KUKA KRL program: folge11.src, folge11.dat

--- folge11.src ---
&ACCESS RVP
&REL 1
&COMMENT bt2krl vw-ks24 production Folge 11 plan 16#F77E
DEF FOLGE11()
   ; Generated by bt2krl 0.1.0 from bt2plc plan bt_1790934549_welding_cell_2_small (cell welding_cell_2_small), PLAN_ID 16#F77E
   ; Robot robot1 (R1), controller 000001R01, model KR240R2900_ULTRA, joint mapping identity
   ; Profile vw-ks24 (VW KS24 / TPVW 8.1.8).
   ; Do not edit: regenerate with bt2krl (plain KRL, no inline forms).
   ; Production Folge: 8 ops; per op: op index BT_PKTNR, interlock request + MAKRO20 handshake, motion (exact stop at the end), hold, interlock release
   ; The VW tech package does the Folge handshake (cell.src, AUE_INIT/WAIT/END).
   ;FOLD AUE INIT
      VW(#VW_AUE_INIT,TRUE)
      PENTER:
      INTERRUPT DECL 10 WHEN $CYCFLAG[254]==FALSE DO VW(#FB_STOP,TRUE)
      INTERRUPT ON 10
      INT10=TRUE
   ;ENDFOLD
   ;FOLD VWP0 P0 10 PCT
      ; P0 = home: VW_INIT runs BAS(#INITMOV); AUE_WAIT later sets $H_POS here
      VW(#VW_INIT,TRUE)
      VW_USR_R (#USR_INIT)
      BAS(#VEL_PTP,10)
      $APO.CPTP=100
      PTP P0
      $OUT[15]=TRUE ; PF0 Grundstellung
      ; MAKRO0 RUECKSETZEN_EA: resets A33-A96 (also the tool releases)
      SEL_RES=SELECT(#MAKRO,0,TRUE,,,,,FALSE)
   ;ENDFOLD
   ;FOLD VWAUEWAIT
      VW(#VW_AUE_WAIT,TRUE )
      IF N_VW==TRUE THEN
         GOTO PEXIT
      ENDIF
   ;ENDFOLD
   ;FOLD VWSTART 16#00000003
      ; release every interlock this robot uses: IL01=V1 IL02=V11
      $OUT[15]=FALSE ; PF0 off
      ; MAKRO50 Ini Merker: the cyclic flags of the driving conditions
      SEL_RES=SELECT(#MAKRO,50,TRUE,,,,,FALSE)
      $OUT[41]=TRUE ; release V1
      $OUT[51]=TRUE ; release V11
   ;ENDFOLD
   ;FOLD PLAN ID 16#F77E
      IF BT_PLANID<>PLAN_ID THEN
         $LOOP_MSG[]="BT2KRL PLAN_ID mismatch - regenerate KRL and PLC"
         HALT
      ENDIF
   ;ENDFOLD
   ;FOLD VWFB 16#00000000
      VALCYCFL30=$CYCFLAG[254]
      $CYCFLAG[254]=($CYCFLAG[30]) AND $CYCFLAG[255] OR ($TIMER[61]<0)
      VW(#FB_CHECK,TRUE)
   ;ENDFOLD
   ;FOLD OP 1 W01 MASK 16#00000001
      ; zones IL01
      BT_PKTNR=1
      ;FOLD VWLOCK 16#00000001
         ; enter IL01=V1
         $OUT[81]=TRUE ; request V1
         ; MAKRO20 semantics, inline for these interlocks only
         $OUT[41]=$OUT[41] OR $OUT[81]
         ; PLC grant of the request
         $LOOP_MSG[]="E81"
         $LOOP_CONT=TRUE
         WAIT FOR ($IN[81]) OR (NOT $LOOP_CONT AND ($MODE_OP<>#EX))
         $LOOP_MSG[]="                                                                                                                                "
         ; partner release
         $LOOP_MSG[]="E41"
         $LOOP_CONT=TRUE
         WAIT FOR ($IN[41]) OR (NOT $LOOP_CONT AND ($MODE_OP<>#EX))
         $LOOP_MSG[]="                                                                                                                                "
         $OUT[41]=FALSE ; occupied
         $OUT[81]=FALSE
      ;ENDFOLD
      ;FOLD VWFB 16#00000001
         VALCYCFL30=$CYCFLAG[254]
         $CYCFLAG[254]=($CYCFLAG[30] AND $IN[41]) AND $CYCFLAG[255] OR ($TIMER[61]<0)
         VW(#FB_CHECK,TRUE)
      ;ENDFOLD
      BAS(#VEL_PTP,3)
      PTP P1 C_PTP
      BAS(#VEL_PTP,6)
      PTP P2 C_PTP
      BAS(#VEL_PTP,10)
      PTP P3 C_PTP
      BAS(#VEL_PTP,12)
      PTP P4 C_PTP
      BAS(#VEL_PTP,15)
      PTP P5 C_PTP
      BAS(#VEL_PTP,17)
      PTP P6 C_PTP
      BAS(#VEL_PTP,19)
      PTP P7 C_PTP
      BAS(#VEL_PTP,17)
      PTP P8 C_PTP
      BAS(#VEL_PTP,13)
      PTP P9 C_PTP
      BAS(#VEL_PTP,10)
      PTP P10 C_PTP
      BAS(#VEL_PTP,6)
      PTP P11 C_PTP
      BAS(#VEL_PTP,3)
      PTP P12 C_PTP
      BAS(#VEL_PTP,5)
      PTP P13 C_PTP
      BAS(#VEL_PTP,4)
      PTP P14
      WAIT SEC 0.5 ; hold
      ;FOLD VWUNLOCK 16#00000001
         ; leave IL01=V1
         $OUT[41]=TRUE ; release V1
      ;ENDFOLD
      ;FOLD VWFB 16#00000000
         VALCYCFL30=$CYCFLAG[254]
         $CYCFLAG[254]=($CYCFLAG[30]) AND $CYCFLAG[255] OR ($TIMER[61]<0)
         VW(#FB_CHECK,TRUE)
      ;ENDFOLD
      WAIT SEC 0.1 ; step dwell
   ;ENDFOLD
   ;FOLD OP 2 W02 MASK 16#00000002
      ; zones IL02
      BT_PKTNR=2
      ;FOLD VWLOCK 16#00000002
         ; enter IL02=V11
         $OUT[91]=TRUE ; request V11
         ; MAKRO20 semantics, inline for these interlocks only
         $OUT[51]=$OUT[51] OR $OUT[91]
         ; PLC grant of the request
         $LOOP_MSG[]="E91"
         $LOOP_CONT=TRUE
         WAIT FOR ($IN[91]) OR (NOT $LOOP_CONT AND ($MODE_OP<>#EX))
         $LOOP_MSG[]="                                                                                                                                "
         ; partner release
         $LOOP_MSG[]="E51"
         $LOOP_CONT=TRUE
         WAIT FOR ($IN[51]) OR (NOT $LOOP_CONT AND ($MODE_OP<>#EX))
         $LOOP_MSG[]="                                                                                                                                "
         $OUT[51]=FALSE ; occupied
         $OUT[91]=FALSE
      ;ENDFOLD
      ;FOLD VWFB 16#00000002
         VALCYCFL30=$CYCFLAG[254]
         $CYCFLAG[254]=($CYCFLAG[30] AND $IN[51]) AND $CYCFLAG[255] OR ($TIMER[61]<0)
         VW(#FB_CHECK,TRUE)
      ;ENDFOLD
      BAS(#VEL_PTP,3)
      PTP P15 C_PTP
      BAS(#VEL_PTP,7)
      PTP P16 C_PTP
      BAS(#VEL_PTP,10)
      PTP P17 C_PTP
      BAS(#VEL_PTP,13)
      PTP P18 C_PTP
      BAS(#VEL_PTP,10)
      PTP P19 C_PTP
      BAS(#VEL_PTP,7)
      PTP P20 C_PTP
      BAS(#VEL_PTP,3)
      PTP P21 C_PTP
      BAS(#VEL_PTP,5)
      PTP P22 C_PTP
      BAS(#VEL_PTP,4)
      PTP P23
      WAIT SEC 0.5 ; hold
      ;FOLD VWUNLOCK 16#00000002
         ; leave IL02=V11
         $OUT[51]=TRUE ; release V11
      ;ENDFOLD
      ;FOLD VWFB 16#00000000
         VALCYCFL30=$CYCFLAG[254]
         $CYCFLAG[254]=($CYCFLAG[30]) AND $CYCFLAG[255] OR ($TIMER[61]<0)
         VW(#FB_CHECK,TRUE)
      ;ENDFOLD
      WAIT SEC 0.1 ; step dwell
   ;ENDFOLD
   ;FOLD OP 3 W03 MASK 16#00000001
      ; zones IL01
      BT_PKTNR=3
      ;FOLD VWLOCK 16#00000001
         ; enter IL01=V1
         $OUT[81]=TRUE ; request V1
         ; MAKRO20 semantics, inline for these interlocks only
         $OUT[41]=$OUT[41] OR $OUT[81]
         ; PLC grant of the request
         $LOOP_MSG[]="E81"
         $LOOP_CONT=TRUE
         WAIT FOR ($IN[81]) OR (NOT $LOOP_CONT AND ($MODE_OP<>#EX))
         $LOOP_MSG[]="                                                                                                                                "
         ; partner release
         $LOOP_MSG[]="E41"
         $LOOP_CONT=TRUE
         WAIT FOR ($IN[41]) OR (NOT $LOOP_CONT AND ($MODE_OP<>#EX))
         $LOOP_MSG[]="                                                                                                                                "
         $OUT[41]=FALSE ; occupied
         $OUT[81]=FALSE
      ;ENDFOLD
      ;FOLD VWFB 16#00000001
         VALCYCFL30=$CYCFLAG[254]
         $CYCFLAG[254]=($CYCFLAG[30] AND $IN[41]) AND $CYCFLAG[255] OR ($TIMER[61]<0)
         VW(#FB_CHECK,TRUE)
      ;ENDFOLD
      BAS(#VEL_PTP,2)
      PTP P24 C_PTP
      BAS(#VEL_PTP,6)
      PTP P25 C_PTP
      BAS(#VEL_PTP,9)
      PTP P26 C_PTP
      BAS(#VEL_PTP,13)
      PTP P27 C_PTP
      BAS(#VEL_PTP,15)
      PTP P28 C_PTP
      BAS(#VEL_PTP,12)
      PTP P29 C_PTP
      BAS(#VEL_PTP,8)
      PTP P30 C_PTP
      BAS(#VEL_PTP,6)
      PTP P31 C_PTP
      BAS(#VEL_PTP,2)
      PTP P32 C_PTP
      BAS(#VEL_PTP,6)
      PTP P33 C_PTP
      BAS(#VEL_PTP,8)
      PTP P34 C_PTP
      BAS(#VEL_PTP,4)
      PTP P35
      WAIT SEC 0.5 ; hold
      ;FOLD VWUNLOCK 16#00000001
         ; leave IL01=V1
         $OUT[41]=TRUE ; release V1
      ;ENDFOLD
      ;FOLD VWFB 16#00000000
         VALCYCFL30=$CYCFLAG[254]
         $CYCFLAG[254]=($CYCFLAG[30]) AND $CYCFLAG[255] OR ($TIMER[61]<0)
         VW(#FB_CHECK,TRUE)
      ;ENDFOLD
      WAIT SEC 0.1 ; step dwell
   ;ENDFOLD
   ;FOLD OP 4 W06 MASK 16#00000002
      ; zones IL02
      BT_PKTNR=4
      ;FOLD VWLOCK 16#00000002
         ; enter IL02=V11
         $OUT[91]=TRUE ; request V11
         ; MAKRO20 semantics, inline for these interlocks only
         $OUT[51]=$OUT[51] OR $OUT[91]
         ; PLC grant of the request
         $LOOP_MSG[]="E91"
         $LOOP_CONT=TRUE
         WAIT FOR ($IN[91]) OR (NOT $LOOP_CONT AND ($MODE_OP<>#EX))
         $LOOP_MSG[]="                                                                                                                                "
         ; partner release
         $LOOP_MSG[]="E51"
         $LOOP_CONT=TRUE
         WAIT FOR ($IN[51]) OR (NOT $LOOP_CONT AND ($MODE_OP<>#EX))
         $LOOP_MSG[]="                                                                                                                                "
         $OUT[51]=FALSE ; occupied
         $OUT[91]=FALSE
      ;ENDFOLD
      ;FOLD VWFB 16#00000002
         VALCYCFL30=$CYCFLAG[254]
         $CYCFLAG[254]=($CYCFLAG[30] AND $IN[51]) AND $CYCFLAG[255] OR ($TIMER[61]<0)
         VW(#FB_CHECK,TRUE)
      ;ENDFOLD
      BAS(#VEL_PTP,8)
      PTP P36 C_PTP
      BAS(#VEL_PTP,16)
      PTP P37 C_PTP
      BAS(#VEL_PTP,8)
      PTP P38 C_PTP
      BAS(#VEL_PTP,4)
      PTP P39 C_PTP
      BAS(#VEL_PTP,3)
      PTP P40
      WAIT SEC 0.5 ; hold
      ;FOLD VWUNLOCK 16#00000002
         ; leave IL02=V11
         $OUT[51]=TRUE ; release V11
      ;ENDFOLD
      ;FOLD VWFB 16#00000000
         VALCYCFL30=$CYCFLAG[254]
         $CYCFLAG[254]=($CYCFLAG[30]) AND $CYCFLAG[255] OR ($TIMER[61]<0)
         VW(#FB_CHECK,TRUE)
      ;ENDFOLD
      WAIT SEC 0.1 ; step dwell
   ;ENDFOLD
   ;FOLD OP 5 W05 MASK 16#00000001
      ; zones IL01
      BT_PKTNR=5
      ;FOLD VWLOCK 16#00000001
         ; enter IL01=V1
         $OUT[81]=TRUE ; request V1
         ; MAKRO20 semantics, inline for these interlocks only
         $OUT[41]=$OUT[41] OR $OUT[81]
         ; PLC grant of the request
         $LOOP_MSG[]="E81"
         $LOOP_CONT=TRUE
         WAIT FOR ($IN[81]) OR (NOT $LOOP_CONT AND ($MODE_OP<>#EX))
         $LOOP_MSG[]="                                                                                                                                "
         ; partner release
         $LOOP_MSG[]="E41"
         $LOOP_CONT=TRUE
         WAIT FOR ($IN[41]) OR (NOT $LOOP_CONT AND ($MODE_OP<>#EX))
         $LOOP_MSG[]="                                                                                                                                "
         $OUT[41]=FALSE ; occupied
         $OUT[81]=FALSE
      ;ENDFOLD
      ;FOLD VWFB 16#00000001
         VALCYCFL30=$CYCFLAG[254]
         $CYCFLAG[254]=($CYCFLAG[30] AND $IN[41]) AND $CYCFLAG[255] OR ($TIMER[61]<0)
         VW(#FB_CHECK,TRUE)
      ;ENDFOLD
      BAS(#VEL_PTP,2)
      PTP P41 C_PTP
      BAS(#VEL_PTP,6)
      PTP P42 C_PTP
      BAS(#VEL_PTP,10)
      PTP P43 C_PTP
      BAS(#VEL_PTP,13)
      PTP P44 C_PTP
      BAS(#VEL_PTP,15)
      PTP P45 C_PTP
      BAS(#VEL_PTP,12)
      PTP P46 C_PTP
      BAS(#VEL_PTP,8)
      PTP P47 C_PTP
      BAS(#VEL_PTP,6)
      PTP P48 C_PTP
      BAS(#VEL_PTP,2)
      PTP P49 C_PTP
      BAS(#VEL_PTP,4)
      PTP P50 C_PTP
      PTP P51
      WAIT SEC 0.5 ; hold
      ;FOLD VWUNLOCK 16#00000001
         ; leave IL01=V1
         $OUT[41]=TRUE ; release V1
      ;ENDFOLD
      ;FOLD VWFB 16#00000000
         VALCYCFL30=$CYCFLAG[254]
         $CYCFLAG[254]=($CYCFLAG[30]) AND $CYCFLAG[255] OR ($TIMER[61]<0)
         VW(#FB_CHECK,TRUE)
      ;ENDFOLD
      WAIT SEC 0.1 ; step dwell
   ;ENDFOLD
   ;FOLD OP 6 W04 MASK 16#00000002
      ; zones IL02
      BT_PKTNR=6
      ;FOLD VWLOCK 16#00000002
         ; enter IL02=V11
         $OUT[91]=TRUE ; request V11
         ; MAKRO20 semantics, inline for these interlocks only
         $OUT[51]=$OUT[51] OR $OUT[91]
         ; PLC grant of the request
         $LOOP_MSG[]="E91"
         $LOOP_CONT=TRUE
         WAIT FOR ($IN[91]) OR (NOT $LOOP_CONT AND ($MODE_OP<>#EX))
         $LOOP_MSG[]="                                                                                                                                "
         ; partner release
         $LOOP_MSG[]="E51"
         $LOOP_CONT=TRUE
         WAIT FOR ($IN[51]) OR (NOT $LOOP_CONT AND ($MODE_OP<>#EX))
         $LOOP_MSG[]="                                                                                                                                "
         $OUT[51]=FALSE ; occupied
         $OUT[91]=FALSE
      ;ENDFOLD
      ;FOLD VWFB 16#00000002
         VALCYCFL30=$CYCFLAG[254]
         $CYCFLAG[254]=($CYCFLAG[30] AND $IN[51]) AND $CYCFLAG[255] OR ($TIMER[61]<0)
         VW(#FB_CHECK,TRUE)
      ;ENDFOLD
      BAS(#VEL_PTP,3)
      PTP P52 C_PTP
      BAS(#VEL_PTP,7)
      PTP P53 C_PTP
      BAS(#VEL_PTP,10)
      PTP P54 C_PTP
      BAS(#VEL_PTP,13)
      PTP P55 C_PTP
      BAS(#VEL_PTP,11)
      PTP P56 C_PTP
      BAS(#VEL_PTP,7)
      PTP P57 C_PTP
      BAS(#VEL_PTP,3)
      PTP P58 C_PTP
      BAS(#VEL_PTP,4)
      PTP P59 C_PTP
      BAS(#VEL_PTP,3)
      PTP P60
      WAIT SEC 0.5 ; hold
      ;FOLD VWUNLOCK 16#00000002
         ; leave IL02=V11
         $OUT[51]=TRUE ; release V11
      ;ENDFOLD
      ;FOLD VWFB 16#00000000
         VALCYCFL30=$CYCFLAG[254]
         $CYCFLAG[254]=($CYCFLAG[30]) AND $CYCFLAG[255] OR ($TIMER[61]<0)
         VW(#FB_CHECK,TRUE)
      ;ENDFOLD
      WAIT SEC 0.1 ; step dwell
   ;ENDFOLD
   ;FOLD OP 7 R1_PARK MASK 16#00000001
      ; zones IL01
      BT_PKTNR=7
      ;FOLD VWLOCK 16#00000001
         ; enter IL01=V1
         $OUT[81]=TRUE ; request V1
         ; MAKRO20 semantics, inline for these interlocks only
         $OUT[41]=$OUT[41] OR $OUT[81]
         ; PLC grant of the request
         $LOOP_MSG[]="E81"
         $LOOP_CONT=TRUE
         WAIT FOR ($IN[81]) OR (NOT $LOOP_CONT AND ($MODE_OP<>#EX))
         $LOOP_MSG[]="                                                                                                                                "
         ; partner release
         $LOOP_MSG[]="E41"
         $LOOP_CONT=TRUE
         WAIT FOR ($IN[41]) OR (NOT $LOOP_CONT AND ($MODE_OP<>#EX))
         $LOOP_MSG[]="                                                                                                                                "
         $OUT[41]=FALSE ; occupied
         $OUT[81]=FALSE
      ;ENDFOLD
      ;FOLD VWFB 16#00000001
         VALCYCFL30=$CYCFLAG[254]
         $CYCFLAG[254]=($CYCFLAG[30] AND $IN[41]) AND $CYCFLAG[255] OR ($TIMER[61]<0)
         VW(#FB_CHECK,TRUE)
      ;ENDFOLD
      BAS(#VEL_PTP,6)
      PTP P61 C_PTP
      BAS(#VEL_PTP,14)
      PTP P62 C_PTP
      BAS(#VEL_PTP,22)
      PTP P63 C_PTP
      BAS(#VEL_PTP,19)
      PTP P64 C_PTP
      BAS(#VEL_PTP,13)
      PTP P65 C_PTP
      BAS(#VEL_PTP,25)
      PTP P66 C_PTP
      PTP P67
      WAIT SEC 0.5 ; hold
      ;FOLD VWUNLOCK 16#00000001
         ; leave IL01=V1
         $OUT[41]=TRUE ; release V1
      ;ENDFOLD
      ;FOLD VWFB 16#00000000
         VALCYCFL30=$CYCFLAG[254]
         $CYCFLAG[254]=($CYCFLAG[30]) AND $CYCFLAG[255] OR ($TIMER[61]<0)
         VW(#FB_CHECK,TRUE)
      ;ENDFOLD
      WAIT SEC 0.1 ; step dwell
   ;ENDFOLD
   ;FOLD OP 8 HOME MASK 16#00000002
      ; zones IL02
      BT_PKTNR=8
      ;FOLD VWLOCK 16#00000002
         ; enter IL02=V11
         $OUT[91]=TRUE ; request V11
         ; MAKRO20 semantics, inline for these interlocks only
         $OUT[51]=$OUT[51] OR $OUT[91]
         ; PLC grant of the request
         $LOOP_MSG[]="E91"
         $LOOP_CONT=TRUE
         WAIT FOR ($IN[91]) OR (NOT $LOOP_CONT AND ($MODE_OP<>#EX))
         $LOOP_MSG[]="                                                                                                                                "
         ; partner release
         $LOOP_MSG[]="E51"
         $LOOP_CONT=TRUE
         WAIT FOR ($IN[51]) OR (NOT $LOOP_CONT AND ($MODE_OP<>#EX))
         $LOOP_MSG[]="                                                                                                                                "
         $OUT[51]=FALSE ; occupied
         $OUT[91]=FALSE
      ;ENDFOLD
      ;FOLD VWFB 16#00000002
         VALCYCFL30=$CYCFLAG[254]
         $CYCFLAG[254]=($CYCFLAG[30] AND $IN[51]) AND $CYCFLAG[255] OR ($TIMER[61]<0)
         VW(#FB_CHECK,TRUE)
      ;ENDFOLD
      BAS(#VEL_PTP,3)
      PTP P68 C_PTP
      BAS(#VEL_PTP,8)
      PTP P69 C_PTP
      BAS(#VEL_PTP,12)
      PTP P70 C_PTP
      BAS(#VEL_PTP,17)
      PTP P71 C_PTP
      BAS(#VEL_PTP,20)
      PTP P72 C_PTP
      BAS(#VEL_PTP,23)
      PTP P73 C_PTP
      BAS(#VEL_PTP,26)
      PTP P74 C_PTP
      BAS(#VEL_PTP,27)
      PTP P75 C_PTP
      BAS(#VEL_PTP,24)
      PTP P76 C_PTP
      BAS(#VEL_PTP,22)
      PTP P77 C_PTP
      BAS(#VEL_PTP,18)
      PTP P78 C_PTP
      BAS(#VEL_PTP,14)
      PTP P79 C_PTP
      BAS(#VEL_PTP,9)
      PTP P80 C_PTP
      BAS(#VEL_PTP,3)
      PTP P81
      ;FOLD VWMAKRO 15
         ; Gesamtfertigmeldung
         SEL_RES=SELECT(#MAKRO,15,TRUE,,,,,FALSE)
      ;ENDFOLD
      ;FOLD VWUNLOCK 16#00000002
         ; leave IL02=V11
         $OUT[51]=TRUE ; release V11
      ;ENDFOLD
      ;FOLD VWFB 16#00000000
         VALCYCFL30=$CYCFLAG[254]
         $CYCFLAG[254]=($CYCFLAG[30]) AND $CYCFLAG[255] OR ($TIMER[61]<0)
         VW(#FB_CHECK,TRUE)
      ;ENDFOLD
      WAIT SEC 0.1 ; step dwell
   ;ENDFOLD
   BT_PKTNR=0
   ;FOLD AUE END
      VW(#VW_AUE_END,TRUE)
      GOTO PENTER
      PEXIT:
   ;ENDFOLD
END

--- folge11.dat ---
&ACCESS RVP
&REL 1
&COMMENT bt2krl vw-ks24 data Folge 11 plan 16#F77E
DEFDAT FOLGE11
   ; Generated by bt2krl 0.1.0 from bt2plc plan bt_1790934549_welding_cell_2_small (cell welding_cell_2_small), PLAN_ID 16#F77E
   ; Robot robot1 (R1), controller 000001R01, model KR240R2900_ULTRA, joint mapping identity
   ; Profile vw-ks24 (VW KS24 / TPVW 8.1.8).
   ; Do not edit: regenerate with bt2krl (plain KRL, no inline forms).
   EXT BAS (BAS_COMMAND :IN,REAL :IN )
   ; interface to the VW standard routines (as every VW Folge .dat declares them)
   EXT VW (VW_COMMAND :IN,BOOL :IN,REAL :IN,REAL :IN,REAL :IN,REAL :IN,BOOL :IN,E6POS :IN )
   EXT VW_USR_R (VW_USER_CMD :IN,INT :IN,REAL :IN,REAL :IN,REAL :IN,REAL :IN,REAL :IN,REAL :IN,BOOL :IN )
   EXTFCT INT SELECT (SUBTYPE :IN,INT :IN,BOOL :IN,ARI_TYP :IN,INT :IN,BOOL_TYP :IN,INT :IN,BOOL :IN)
   DECL AXIS P0={A1 0.0,A2 -90.0,A3 90.0,A4 0.0,A5 0.0,A6 0.0}
   DECL AXIS P1={A1 -1.1481,A2 -89.8273,A3 90.1392,A4 0.2955,A5 0.7752,A6 0.3515}
   DECL AXIS P2={A1 -4.4157,A2 -89.3356,A3 90.5354,A4 1.1366,A5 2.9817,A6 1.3518}
   DECL AXIS P3={A1 -9.5379,A2 -88.565,A3 91.1564,A4 2.455,A5 6.4405,A6 2.9199}
   DECL AXIS P4={A1 -16.2497,A2 -87.5551,A3 91.9702,A4 4.1827,A5 10.9727,A6 4.9746}
   DECL AXIS P5={A1 -24.2863,A2 -86.346,A3 92.9446,A4 6.2512,A5 16.3994,A6 7.4349}
   DECL AXIS P6={A1 -38.2454,A2 -84.2458,A3 94.6371,A4 9.8443,A5 25.8253,A6 11.7083}
   DECL AXIS P7={A1 -90.5161,A2 -76.3814,A3 100.9747,A4 23.2987,A5 61.1212,A6 27.7103}
   DECL AXIS P8={A1 -108.6425,A2 -73.6542,A3 103.1724,A4 27.9644,A5 73.3611,A6 33.2594}
   DECL AXIS P9={A1 -119.2236,A2 -72.0622,A3 104.4553,A4 30.6879,A5 80.506,A6 36.4987}
   DECL AXIS P10={A1 -124.3458,A2 -71.2916,A3 105.0764,A4 32.0064,A5 83.9648,A6 38.0668}
   DECL AXIS P11={A1 -127.6134,A2 -70.7999,A3 105.4725,A4 32.8474,A5 86.1712,A6 39.0671}
   DECL AXIS P12={A1 -128.7615,A2 -70.6272,A3 105.6117,A4 33.143,A5 86.9465,A6 39.4186}
   DECL AXIS P13={A1 -128.7615,A2 -70.2228,A3 105.9156,A4 33.18,A5 86.8872,A6 39.3731}
   DECL AXIS P14={A1 -128.7615,A2 -67.4517,A3 107.7396,A4 33.6697,A5 83.7898,A6 37.2493}
   DECL AXIS P15={A1 -128.6426,A2 -67.6366,A3 107.8186,A4 32.7502,A5 82.9536,A6 37.7433}
   DECL AXIS P16={A1 -128.3199,A2 -68.1386,A3 108.0329,A4 30.2544,A5 80.6837,A6 39.084}
   DECL AXIS P17={A1 -127.8443,A2 -68.8784,A3 108.3488,A4 26.5764,A5 77.3387,A6 41.0597}
   DECL AXIS P18={A1 -125.4325,A2 -72.6301,A3 109.9508,A4 7.9238,A5 60.3747,A6 51.0796}
   DECL AXIS P19={A1 -124.957,A2 -73.3699,A3 110.2667,A4 4.2458,A5 57.0297,A6 53.0553}
   DECL AXIS P20={A1 -124.6342,A2 -73.8718,A3 110.481,A4 1.75,A5 54.7598,A6 54.396}
   DECL AXIS P21={A1 -124.5154,A2 -74.0568,A3 110.56,A4 0.8305,A5 53.9236,A6 54.8899}
   DECL AXIS P22={A1 -124.5151,A2 -73.6213,A3 110.8768,A4 0.5687,A5 53.3206,A6 55.0767}
   DECL AXIS P23={A1 -124.5148,A2 -70.6583,A3 112.7632,A4 0.0121,A5 48.729,A6 55.4761}
   DECL AXIS P24={A1 -124.4617,A2 -70.7313,A3 112.7862,A4 -0.6572,A5 48.6812,A6 55.9965}
   DECL AXIS P25={A1 -124.3117,A2 -70.9378,A3 112.8512,A4 -2.5487,A5 48.5461,A6 57.4671}
   DECL AXIS P26={A1 -123.7762,A2 -71.6746,A3 113.0835,A4 -9.2998,A5 48.0639,A6 62.7161}
   DECL AXIS P27={A1 -123.0192,A2 -72.7163,A3 113.4118,A4 -18.8444,A5 47.3821,A6 70.1371}
   DECL AXIS P28={A1 -120.8842,A2 -75.654,A3 114.3378,A4 -45.7616,A5 45.4595,A6 91.0652}
   DECL AXIS P29={A1 -120.2241,A2 -76.5623,A3 114.6241,A4 -54.084,A5 44.865,A6 97.536}
   DECL AXIS P30={A1 -119.991,A2 -76.883,A3 114.7252,A4 -57.0231,A5 44.6551,A6 99.8211}
   DECL AXIS P31={A1 -119.8409,A2 -77.0895,A3 114.7902,A4 -58.9146,A5 44.52,A6 101.2917}
   DECL AXIS P32={A1 -119.7879,A2 -77.1625,A3 114.8133,A4 -59.5839,A5 44.4722,A6 101.8121}
   DECL AXIS P33={A1 -119.7876,A2 -76.7001,A3 115.1416,A4 -60.3559,A5 44.324,A6 102.6809}
   DECL AXIS P34={A1 -119.7872,A2 -76.0201,A3 115.6192,A4 -61.4852,A5 44.0795,A6 103.9753}
   DECL AXIS P35={A1 -119.7872,A2 -73.5459,A3 117.1,A4 -65.4365,A5 42.4249,A6 109.2463}
   DECL AXIS P36={A1 -119.1489,A2 -72.8001,A3 114.8711,A4 -64.2164,A5 43.4199,A6 108.0229}
   DECL AXIS P37={A1 -116.34,A2 -69.5185,A3 105.0638,A4 -58.8479,A5 47.7981,A6 102.6395}
   DECL AXIS P38={A1 -115.7016,A2 -68.7727,A3 102.8349,A4 -57.6278,A5 48.7931,A6 101.416}
   DECL AXIS P39={A1 -115.7012,A2 -68.3831,A3 103.1319,A4 -57.6419,A5 48.7925,A6 101.457}
   DECL AXIS P40={A1 -115.7007,A2 -65.7101,A3 104.9261,A4 -60.3105,A5 47.1665,A6 105.7542}
   DECL AXIS P41={A1 -115.7494,A2 -65.7146,A3 104.8564,A4 -59.6416,A5 47.2762,A6 105.2455}
   DECL AXIS P42={A1 -115.887,A2 -65.727,A3 104.6592,A4 -57.7513,A5 47.5859,A6 103.8079}
   DECL AXIS P43={A1 -116.378,A2 -65.7715,A3 103.9556,A4 -51.0043,A5 48.6915,A6 98.6766}
   DECL AXIS P44={A1 -117.0722,A2 -65.8345,A3 102.9609,A4 -41.4655,A5 50.2545,A6 91.4221}
   DECL AXIS P45={A1 -119.0301,A2 -66.012,A3 100.1555,A4 -14.5649,A5 54.6625,A6 70.9633}
   DECL AXIS P46={A1 -119.6354,A2 -66.0668,A3 99.2881,A4 -6.2475,A5 56.0254,A6 64.6377}
   DECL AXIS P47={A1 -119.8492,A2 -66.0862,A3 98.9818,A4 -3.3103,A5 56.5068,A6 62.4038}
   DECL AXIS P48={A1 -119.9868,A2 -66.0987,A3 98.7847,A4 -1.42,A5 56.8165,A6 60.9662}
   DECL AXIS P49={A1 -120.0355,A2 -66.1031,A3 98.7149,A4 -0.7511,A5 56.9261,A6 60.4575}
   DECL AXIS P50={A1 -120.0357,A2 -65.7312,A3 99.0104,A4 -0.6308,A5 56.7548,A6 60.3791}
   DECL AXIS P51={A1 -120.0359,A2 -63.1985,A3 100.772,A4 -0.0303,A5 53.2125,A6 59.9847}
   DECL AXIS P52={A1 -120.1288,A2 -63.1954,A3 100.6111,A4 0.7952,A5 54.0248,A6 59.6456}
   DECL AXIS P53={A1 -120.3834,A2 -63.1866,A3 100.1699,A4 3.0584,A5 56.2523,A6 58.7158}
   DECL AXIS P54={A1 -120.7638,A2 -63.1736,A3 99.5107,A4 6.44,A5 59.5803,A6 57.3266}
   DECL AXIS P55={A1 -122.8245,A2 -63.1028,A3 95.9394,A4 24.7593,A5 77.6095,A6 49.8008}
   DECL AXIS P56={A1 -123.6751,A2 -63.0736,A3 94.4653,A4 32.3213,A5 85.0518,A6 46.6942}
   DECL AXIS P57={A1 -123.9297,A2 -63.0649,A3 94.024,A4 34.5845,A5 87.2792,A6 45.7644}
   DECL AXIS P58={A1 -124.0225,A2 -63.0617,A3 93.8631,A4 35.41,A5 88.0916,A6 45.4253}
   DECL AXIS P59={A1 -124.0227,A2 -62.712,A3 94.1541,A4 35.4756,A5 88.0225,A6 45.3131}
   DECL AXIS P60={A1 -124.0229,A2 -60.325,A3 95.8907,A4 35.9822,A5 85.4859,A6 43.0775}
   DECL AXIS P61={A1 -125.6247,A2 -60.4541,A3 95.8014,A4 35.9822,A5 85.4859,A6 43.0775}
   DECL AXIS P62={A1 -129.8294,A2 -60.7871,A3 95.5713,A4 35.9822,A5 85.4859,A6 43.0775}
   DECL AXIS P63={A1 -149.0509,A2 -62.195,A3 94.602,A4 35.9822,A5 85.4859,A6 43.0775}
   DECL AXIS P64={A1 -154.6572,A2 -62.529,A3 94.3745,A4 35.9822,A5 85.4859,A6 43.0775}
   DECL AXIS P65={A1 -158.3613,A2 -62.6594,A3 94.2891,A4 35.9822,A5 85.4859,A6 43.0775}
   DECL AXIS P66={A1 -160.5075,A2 -61.5043,A3 95.1253,A4 35.9822,A5 85.4859,A6 43.0775}
   DECL AXIS P67={A1 -158.3613,A2 -60.3464,A3 95.9536,A4 35.9822,A5 85.4859,A6 43.0775}
   DECL AXIS P68={A1 -157.2676,A2 -60.5512,A3 95.9125,A4 35.7336,A5 84.8955,A6 42.78}
   DECL AXIS P69={A1 -154.1335,A2 -61.1381,A3 95.7947,A4 35.0215,A5 83.2037,A6 41.9274}
   DECL AXIS P70={A1 -149.1796,A2 -62.0657,A3 95.6084,A4 33.8959,A5 80.5295,A6 40.5799}
   DECL AXIS P71={A1 -138.8192,A2 -64.0057,A3 95.2189,A4 31.5419,A5 74.9368,A6 37.7616}
   DECL AXIS P72={A1 -130.2809,A2 -65.6046,A3 94.8979,A4 29.6018,A5 70.3276,A6 35.439}
   DECL AXIS P73={A1 -115.5777,A2 -68.3578,A3 94.3452,A4 26.2611,A5 62.3907,A6 31.4395}
   DECL AXIS P74={A1 -99.2616,A2 -71.413,A3 93.7317,A4 22.5538,A5 53.583,A6 27.0012}
   DECL AXIS P75={A1 -48.0798,A2 -80.9969,A3 91.8076,A4 10.9245,A5 25.9542,A6 13.0787}
   DECL AXIS P76={A1 -32.7563,A2 -83.8663,A3 91.2315,A4 7.4427,A5 17.6824,A6 8.9104}
   DECL AXIS P77={A1 -23.6665,A2 -85.5684,A3 90.8897,A4 5.3774,A5 12.7756,A6 6.4378}
   DECL AXIS P78={A1 -12.2721,A2 -87.702,A3 90.4614,A4 2.7884,A5 6.6247,A6 3.3383}
   DECL AXIS P79={A1 -6.4911,A2 -88.7845,A3 90.244,A4 1.4749,A5 3.504,A6 1.7657}
   DECL AXIS P80={A1 -1.0937,A2 -89.7952,A3 90.0411,A4 0.2485,A5 0.5904,A6 0.2975}
   DECL AXIS P81={A1 0.0,A2 -90.0,A3 90.0,A4 0.0,A5 0.0,A6 0.0}
ENDDAT
